(* IEC 61131-3 sources: SortJet_MasterSPS_Aufbau.fbsproj/Device.device.xml.v3^/Plc Logic.plclogic.xml.v3^/Application.application.xml.v3^/09_Station/Shuttle/Zentralschmierung, 1 file *)

(* ---- MK_Zentralschmierung.gvl ---- *)
(* METADATA
{
	"v3Meta": {
		"objectGuid": "cea505f7-1a84-4065-b281-2c700363fb8a"
	}
}
*)
{attribute 'allow_unqualified_access'}
NAMESPACE MK_Zentralschmierung
VAR_GLOBAL

  // Zentralschmierung Shuttle
  apgMKShuttleZentralschmierung : ARRAY [cERSTES_SHUTTLE..cLETZTES_SHUTTLE] OF Parameter_Zentralschmierung_DLS_4xxi :=[
    // ----------------------------------- SHUTTLE 101 ---------------------------------------------------
    (
      aiAnzahlHuebe                   := [3,20],             // Anzahl der Hübe die die Schmierung machen soll
      adiZuFahrenderWegBisSchmierung  := [21600000,24500000] // Zu fahrende Strecke nach der geschmiert werden muss in mm
    ),
    // ----------------------------------- SHUTTLE 102 ---------------------------------------------------
    (
      aiAnzahlHuebe                   := [3,20],             // Anzahl der Hübe die die Schmierung machen soll
      adiZuFahrenderWegBisSchmierung  := [21600000,24500000] // Zu fahrende Strecke nach der geschmiert werden muss in mm
    )];

  // Zentralschmierung Transfershuttle
  apgMKTransfershuttleZentralschmierung : ARRAY [cERSTES_TRANSFERSHUTTLE..cLETZTES_TRANSFERSHUTTLE ] OF Parameter_Zentralschmierung_DLS_4xxi :=[
    // ----------------------------------- TRANSFERSHUTTLE 151 ---------------------------------------------------
    (
      aiAnzahlHuebe                   := [3,20],             // Anzahl der Hübe die die Schmierung machen soll
      adiZuFahrenderWegBisSchmierung  := [11300000,40500000] // Zu fahrende Strecke nach der geschmiert werden muss in mm
    ),
    // ----------------------------------- TRANSFERSHUTTLE 152 ---------------------------------------------------
    (
      aiAnzahlHuebe                   := [3,20],             // Anzahl der Hübe die die Schmierung machen soll
      adiZuFahrenderWegBisSchmierung  := [11300000,40500000] // Zu fahrende Strecke nach der geschmiert werden muss in mm
    )];

END_VAR
END_NAMESPACE
